Fanuc KAREL source: KT00905.KL

PROGRAM KT00905
%NOLOCKGROUP
%ENVIRONMENT VECTR
VAR
  P1: XYZWPREXT
  P2: XYZWPREXT
  OUT: VECTOR
BEGIN
  P1.X = 1.0
  P2.Y = 2.0
  P1.X = 1.0
  P2.Y = 2.0
  OUT = APPROACH(P1)
END KT00905
